(* IEC 61131-3 sources: nautilus/tools/blackbox/projects/2026-10-24-001/mb, 1 file *)

(* ---- main.st ---- *)
PROGRAM Main
VAR_EXTERNAL
    Beat : DINT;
END_VAR
Beat := Beat + 1;
END_PROGRAM
